FUNCTION_BLOCK F_Concat_Tests EXTENDS TcUnit.FB_TestSuite

Test_Concat3();
Test_Concat4();
Test_Concat5();
Test_Concat6();
Test_Concat7();
Test_EmptyPartsAreSkipped();
Test_ResultLimitedToMaxString();

METHOD PRIVATE Test_Concat3
TcUnit.TEST(__POUNAME());

AssertEquals_STRING(Expected := 'abc', Actual := F_Concat3('a', 'b', 'c'), Message := 'three parts joined');

TEST_FINISHED_NAMED(__POUNAME());
END_METHOD

METHOD PRIVATE Test_Concat4
TcUnit.TEST(__POUNAME());

AssertEquals_STRING(Expected := 'abcd', Actual := F_Concat4('a', 'b', 'c', 'd'), Message := 'four parts joined');

TEST_FINISHED_NAMED(__POUNAME());
END_METHOD

METHOD PRIVATE Test_Concat5
TcUnit.TEST(__POUNAME());

AssertEquals_STRING(Expected := 'abcde', Actual := F_Concat5('a', 'b', 'c', 'd', 'e'), Message := 'five parts joined');

TEST_FINISHED_NAMED(__POUNAME());
END_METHOD

METHOD PRIVATE Test_Concat6
TcUnit.TEST(__POUNAME());

AssertEquals_STRING(Expected := 'abcdef', Actual := F_Concat6('a', 'b', 'c', 'd', 'e', 'f'), Message := 'six parts joined');

TEST_FINISHED_NAMED(__POUNAME());
END_METHOD

METHOD PRIVATE Test_Concat7
TcUnit.TEST(__POUNAME());

AssertEquals_STRING(Expected := 'abcdefg', Actual := F_Concat7('a', 'b', 'c', 'd', 'e', 'f', 'g'), Message := 'seven parts joined');

TEST_FINISHED_NAMED(__POUNAME());
END_METHOD

METHOD PRIVATE Test_EmptyPartsAreSkipped
TcUnit.TEST(__POUNAME());

AssertEquals_STRING(Expected := 'x', Actual := F_Concat3('', 'x', ''), Message := 'empty parts contribute nothing');

TEST_FINISHED_NAMED(__POUNAME());
END_METHOD

METHOD PRIVATE Test_ResultLimitedToMaxString
VAR
  part : STRING;
  i : INT;
  result : T_MaxString;
END_VAR
TcUnit.TEST(__POUNAME());

// arrange
FOR i := 1 TO 80 DO
  part := CONCAT(part, 'x');
END_FOR

// act
result := F_Concat4(part, part, part, part);

// assert
AssertEquals_INT(Expected := 255, Actual := LEN(result), Message := '4 x 80 characters truncate to T_MaxString');

TEST_FINISHED_NAMED(__POUNAME());
END_METHOD

END_FUNCTION_BLOCK

(* stored: Version 1.1.0.1, ProductVersion 3.1.4026.22
   POU F_Concat_Tests: Id {d21c9e8d-b8fd-4e4a-b543-1180e84d90a6}, SpecialFunc None
   Method Test_Concat3: Id {2441c1cd-bd4d-44c6-a97f-c8219faf81d1}
   Method Test_Concat4: Id {5eb7d0fd-c52b-4901-a872-3a8507937325}
   Method Test_Concat5: Id {7883ccc4-0d28-4ae2-b09e-287e348d4b43}
   Method Test_Concat6: Id {284ee546-71f7-4740-83e4-3ac8c6281749}
   Method Test_Concat7: Id {6f7ae99e-475f-4863-b29e-b22c36af9eaa}
   Method Test_EmptyPartsAreSkipped: Id {103788f2-9614-472e-8298-a3fee5b01895}
   Method Test_ResultLimitedToMaxString: Id {dc12d384-7b9f-4215-a3fe-95b4a2ac5f92} *)
